// TIA Portal V20 export
// export: Created 2026-10-12T16:46:22.7860407Z, ExportSetting WithDefaults, DisplayName Totally Integrated Automation Portal, DisplayVersion V20 Update 6, DisplayName TIA Portal Openness, DisplayVersion V20 Update 6, DisplayName TIA Portal Version Control Interface, DisplayVersion V20 Update 6, DisplayName SINAMICS Startdrive Advanced, DisplayVersion V20 SP1 Update 2, DisplayName SINAMICS Startdrive G110M, G120, G120C, G120D, G120P, G115D, DisplayVersion V20 SP1 Update 2, DisplayName SINAMICS Startdrive G130, G150, S120, S150, SINAMICS MV, G220, S200, S210, DisplayVersion V20 SP1 Update 2, DisplayName STEP 7 Professional, DisplayVersion V20 Update 6, DisplayName STEP 7 Safety, DisplayVersion V20 Update 2, DisplayName WinCC Basic/Comfort/Advanced, DisplayVersion V20 Update 6, DisplayName WinCC Professional, DisplayVersion V20 Update 6, DisplayName WinCC Unified, DisplayVersion V20 Update 6
TYPE "UDT_Handbetrieb"
// stored: IsFailsafeCompliant false
   STRUCT
      Hand_Aktiv : Bool;
      Pumpe : Bool;
      Pumpe_FU_Soll : Real;   // Umwaelzpumpe Drehzahl (%)
      Ultraschall : Bool;
      Heizung_Soll : Real;
      GR_Aktiv : Bool;
      GR_Strom_Soll : Real;
      GR_Spannung_Soll : Real;
      GR_Pulsfrequenz : Real;
      GR_DutyCycle : Real;
      Warenbewegung_X : Real;
      Warenbewegung_Y : Real;
      WB1_Reset : Bool;   // FU Reset Warenbewegung 1
      WB2_Reset : Bool;   // FU Reset Warenbewegung 2
      Pumpe_FU_Reset : Bool;   // FU Reset Umwaelzpumpe
   END_STRUCT;
END_TYPE
